// TIA Portal V20 export
// export: Created 2026-10-19T18:05:41.00076Z, ExportSetting WithDefaults, DisplayName Totally Integrated Automation Portal, DisplayVersion V20 Update 6, DisplayName TIA Portal Openness, DisplayVersion V20 Update 6, DisplayName TIA Portal Version Control Interface, DisplayVersion V20 Update 6, DisplayName SINAMICS Startdrive Advanced, DisplayVersion V20 SP1, DisplayName SINAMICS Startdrive G130, G150, S120, S150, SINAMICS MV, G220, S200, S210, DisplayVersion V20 SP1, DisplayName SINAMICS Startdrive G110M, G120, G120C, G120D, G120P, G115D, DisplayVersion V20 SP1, DisplayName STEP 7 Professional, DisplayVersion V20 Update 6, DisplayName STEP 7 Safety, DisplayVersion V20 Update 2, DisplayName WinCC Basic/Comfort/Advanced, DisplayVersion V20 Update 6, DisplayName WinCC Unified, DisplayVersion V20 Update 6
FUNCTION "FindBoolField" : Bool   // FC17, SCL
{ S7_Optimized_Access := 'TRUE' }
VERSION : 0.1
// stored: AutoNumber true, IsIECCheckEnabled false, SetENOAutomatically false, UDAEnableTagReadback false
   VAR_INPUT
      FieldName : String;
      JsonStr : String;
   END_VAR
   VAR_TEMP
      searchStr : String;
      foundPos : Int;
      valueStr : String;
      afterField : String;
      bResult : Bool;
   END_VAR
BEGIN
   // Build search string
   #searchStr := CONCAT(IN1 := '"', IN2 := #FieldName);
   #searchStr := CONCAT(IN1 := #searchStr, IN2 := '" :');

   // Serach for JSON field
   #foundPos := FIND(IN1 := #JsonStr, IN2 := #searchStr);

   IF #foundPos > 0 THEN
       // Take to 20 characters after the field
       #afterField := MID(IN := #JsonStr, P := #foundPos + LEN(#searchStr), L := 20);

       // Normalize to remove whitespace if necessary
       // (or compare directly)
       IF FIND(IN1 := #afterField, IN2 := 'true') > 0 THEN
           #bResult := TRUE;
       ELSIF FIND(IN1 := #afterField, IN2 := 'false') > 0 THEN
           #bResult := FALSE;
       ELSE
           #bResult := FALSE; // default if value not found
       END_IF;
   ELSE
       #bResult := FALSE;
   END_IF;

   #FindBoolField := #bResult;
END_FUNCTION
